Fanuc KAREL source: KA00147.KL

PROGRAM KA00147
%NOLOCKGROUP
VAR
  SRC: ARRAY[4] OF INTEGER
  DST: ARRAY[4] OF BOOLEAN
BEGIN
  DST = SRC
END KA00147
